{region 'Documentation'}
(*!
<summary>Checks that IN is a finite value.</summary>
<description>

NaN and either infinity are legitimate checked data, not configuration errors.
Classification mismatch reports Failed. Bit-based classification does not perform an ordered
floating-point comparison.

Numeric diagnostics use the formatter's default six significant digits; rounding affects
the message only, not the comparison.

</description>
*)
{endregion}
FUNCTION_BLOCK AssertIsFinite_LReal EXTENDS AssertionBase
VAR_INPUT
    IN : LREAL; //! Value to classify; NaN and both infinities are valid inputs.
END_VAR

SUPER^();

{region 'Documentation'}
(*!
<summary>Classifies the bit representation without floating-point arithmetic.</summary>
*)
{endregion}
METHOD PROTECTED Assert
VAR
    Representation : AssertionLRealRepresentation;
    Message : STRING(GVL_Constants.MessageLength);
END_VAR
VAR CONSTANT
    ExponentMask : LWORD := LWORD#16#7FF0000000000000;
END_VAR
IF NOT EvaluationActive THEN
    RETURN;
END_IF;

IF Result = E_Result.Error THEN
    RETURN;
END_IF;

IF Result = E_Result.Failed THEN
    RETURN;
END_IF;

Representation.Value := IN;
IF (Representation.Bits AND ExponentMask) = ExponentMask THEN
    Message := CONCAT('Assertion failed: expected a finite value. Actual = ',
        CreateAssertionTextValue_LReal(Value := IN));
    Message := CONCAT(Message, '.');
    Fail(Message := Message);
    RETURN;
END_IF;

Pass();
END_METHOD

END_FUNCTION_BLOCK

(* stored: Version 1.1.0.1
   POU AssertIsFinite_LReal: Id {4cfdd34e-10da-45ed-9842-4c1082cb9379}, SpecialFunc None
   Folder Internal: Id {5291b086-62d9-4419-ab39-7e636565863f}
   Method Assert: Id {a6310000-0000-4000-8000-000000000004} *)
